Fanuc KAREL source: KA00212.KL

PROGRAM KA00212
%NOLOCKGROUP
VAR
  SRC: ARRAY[4] OF XYZWPR
  DST: ARRAY[4] OF BYTE
BEGIN
  DST = SRC
END KA00212
